(* IEC 61131-3 sources: ConveyorControl-with-PLC/4E_Gruppe1_Graf_Projekt1/Class/SafetyBase (part 5) *)

            // get state via SDO communication
            StandardRequest.SDOHeader.CRC  := 0;                                                   // CRC is always 0 in Std communication
            StandardRequest.SDOHeader.Cmd  := SB_SDO_COMMAND_GET_DIAG_INFO;                        // read command
            StandardRequest.SDOHeader.Typ  := SDO_STD;                                             // standard frame type
            StandardRequest.SDOHeader.SeqNr:= StandardSeqNr OR 16#80;                              // sequence number
            StandardRequest.SDOHeader.Len  := 4 + 1;                                               // header + µC-selection
            StandardRequest.aData[0] := DiagVars.ucChoiceDiagInfo;

            LastRequest := _DiagInfo;

#ifdef SAFETY_PROTOCOL_ANALYZER_ACTIVATED
  RecordFrame((#StandardRequest)$^DINT, 1);
#endif

            //copy SDO into write-buffer
            ToStdLib.MemCpy(dest := #p_Handle_SDO_Write^.SDOStructure, source := #StandardRequest, size := (sizeof(SDOHeader.StdHeader.CRC) + StandardRequest.SDOHeader.Len));

            //mark SDO data as valid
            p_Handle_SDO_Write^.us_Status := SAFETY_SDO_DATA_VALID;

            if ( pISafety^.udVersion >= 16#1001 ) then
              SAFETY_iPushSafetyTask();
            end_if;

          else

            if SchedulerStepNo = 6 then
              UnsafeScheduler := UnsafeSchedulerGetDiagVars;

            elsif SchedulerStepNo = 7 then
              UnsafeScheduler := UnsafeSchedulerGetRetryCounter;
            end_if;

          end_if;
       (* ***************************************** *)
          UnsafeSchedulerGetRetryCounter:
       (* ***************************************** *)
           //read out the retry counters every 10seconds
          if (ops.tAbsolute - ud_RetryCntTimeMark) > SB_RETRY_COUNTER_WAIT_TIME  then

            SDORequestBuffer.StdHeader.CRC  := 0;                                                         // CRC is always 0 in Std communication
            SDORequestBuffer.StdHeader.Cmd  := SB_SDO_COMMAND_READ;                                       // read command
            SDORequestBuffer.StdHeader.Typ  := SDO_STD;                                                   // standard frame type
            SDORequestBuffer.StdHeader.SeqNr:= StandardSeqNr OR 16#80;                                    // sequence number
            SDORequestBuffer.StdHeader.Len  := 4 + 4 + SB_SDO_LENGTH_RETRY_COUNTER;                       // header + destination address + length of data
            SDORequestBuffer.ud_Address     := SB_SDO_ADDRESS_RETRY_COUNTER;                              // address of retrycounter
            SDORequestBuffer.us_Length      := SB_SDO_LENGTH_RETRY_COUNTER;                               // length of data

            LastRequest := _ReadRetryCounter;

  #ifdef SAFETY_PROTOCOL_ANALYZER_ACTIVATED
  RecordFrame((#SDORequestBuffer)$^DINT, 1);
  #endif

            //copy SDO into write-buffer
            ToStdLib.MemCpy(dest := #p_Handle_SDO_Write^.SDOStructure, source := #SDORequestBuffer, size := (sizeof(SDOHeader.StdHeader.CRC) + SDORequestBuffer.StdHeader.Len));

            //mark SDO data as valid
            p_Handle_SDO_Write^.us_Status := SAFETY_SDO_DATA_VALID;

            if ( pISafety^.udVersion >= 16#1001 ) then
              SAFETY_iPushSafetyTask();
            end_if;

            //reset timemark
            ud_RetryCntTimeMark := ops.tAbsolute;

          else
            UnsafeScheduler := UnsafeSchedulerGetDiagVars;
          end_if;
        else
          LogError("Undefined Scheduler-State");
        end_case;
      end_while;
    end_if;
  end_if;

  // at the first run we write all variables independent of any changes
  if RunState > OldRunState then
    SendAllUnsafeValues();
  end_if;
  OldRunState := RunState;

	state := READY;

//============================ Profiler start======================================================
#ifdef  DM_Profiler
  StopTimeMeasurement(usMode := DMTIME_CY);
#endif
//============================ Profiler end========================================================
END_FUNCTION

FUNCTION SafetyBase::GetPointer2IFPDOBuffer
	VAR_OUTPUT
		ud_PDOBuffer 	: UDINT;
	END_VAR

  IFPDOOutputIsUsed := TRUE;

  //set pointer to address of buffer pointer
  ud_PDOBuffer := ( #IFPDOOutputBuffer )$UDINT;

END_FUNCTION

FUNCTION VIRTUAL SafetyBase::GetConfiguration

END_FUNCTION

FUNCTION SafetyBase::AddMovDOs
	VAR_OUTPUT
		ret_code 	: iprStates;
	END_VAR
  VAR
  	tempCmd         : CmdStruct;
    _result         : results;
    dataADDDO       : t_AddMoveDOCfg;
    i               : DINT;
  END_VAR

  ret_code := READY;

  // at the connect of the module we read the needed write size (written by the safety designer). at this point we know if the module needs data. if not => no move necessary
  if MyPDOWriteSize = 0 then
    return;
  end_if;

  // this stays the same for every DO
  tempCmd.uiCmd     := _BUS_IF_ADD_MOVE_DO;
  tempCmd.aPara[0]  := (#dataADDDO)$DINT;

  // initialize the parameter structure
  dataADDDO.ud_length_move        := MyPDOWriteSize;
  dataADDDO.ud_handle_source      := 0; // is set via SdiasManager or similar
  dataADDDO.ud_addressoff_source  := 0; // is set via SdiasManager or similar
  dataADDDO.p_sourcedata          := pPDOReadData;
  dataADDDO.ud_handle_dest        := 0; // is set via SdiasManager or similar
  dataADDDO.ud_addressoff_dest    := 0; // is set via SdiasManager or similar
  dataADDDO.p_destdata            := pPDOWriteData;
  dataADDDO.Priority              := _BUS_IF_ISO_MOVE;

  ToBusInterface.NewInst(pPara:=#tempCmd, pResult:=#_result);
  if _result.aData[0]$t_BusIFRetvalErrorcode = _BUS_IF_RETVAL_OK then
    InputMovSettings.MoveSettingsBusIF.Handle               := _result.aData$t_AddMoveDORet.Handle;
    InputMovSettings.MoveSettingsBusIF.ud_length_move       := dataADDDO.ud_length_move;
    InputMovSettings.MoveSettingsBusIF.ud_handle_source     := dataADDDO.ud_handle_source;
    InputMovSettings.MoveSettingsBusIF.ud_addressoff_source := dataADDDO.ud_addressoff_source;
    InputMovSettings.MoveSettingsBusIF.p_sourcedata         := dataADDDO.p_sourcedata;
    InputMovSettings.MoveSettingsBusIF.ud_handle_dest       := dataADDDO.ud_handle_dest;
    InputMovSettings.MoveSettingsBusIF.ud_addressoff_dest   := dataADDDO.ud_addressoff_dest;
    InputMovSettings.MoveSettingsBusIF.p_destdata           := dataADDDO.p_destdata;
    InputMovSettings.EnableState                            := _BUS_IF_RUN_STATE_NO_RUN;

    // addresses of local PDOs (set after creating the Move-DO, because we don't have the pointers to the DPRAM before (only in local memory)
    ud_LocalMoveSourceAddr := dataADDDO.p_sourcedata$UDINT;
    ud_LocalMoveDestAddr   := dataADDDO.p_destdata$UDINT;

    ud_LocalReadHandle     := dataADDDO.ud_handle_source;
    ud_LocalReadOffset     := dataADDDO.ud_addressoff_source;

    ud_LocalWriteHandle    := dataADDDO.ud_handle_dest;
    ud_LocalWriteOffset    := dataADDDO.ud_addressoff_dest;
  else
    LogError("(SafetyBase::AddMovDOs) Failed to add move DO");
    ret_code := ERROR;
  end_if;

  if (AdditionalSPDOs > 0) then
    for i := 0 to (AdditionalSPDOs-1) do
      dataADDDO.p_destdata  := aAdditionalPDOs[i].pPDOWriteData;

      ToBusInterface.NewInst(pPara:=#tempCmd, pResult:=#_result);
      if _result.aData[0]$t_BusIFRetvalErrorcode = _BUS_IF_RETVAL_OK then
        aAdditionalPDOs[i].InputMovSettings.MoveSettingsBusIF.Handle                := _result.aData$t_AddMoveDORet.Handle;
        aAdditionalPDOs[i].InputMovSettings.MoveSettingsBusIF.ud_length_move        := dataADDDO.ud_length_move;
        aAdditionalPDOs[i].InputMovSettings.MoveSettingsBusIF.ud_handle_source      := dataADDDO.ud_handle_source;
        aAdditionalPDOs[i].InputMovSettings.MoveSettingsBusIF.ud_addressoff_source  := dataADDDO.ud_addressoff_source;
        aAdditionalPDOs[i].InputMovSettings.MoveSettingsBusIF.p_sourcedata          := dataADDDO.p_sourcedata;
        aAdditionalPDOs[i].InputMovSettings.MoveSettingsBusIF.ud_handle_dest        := dataADDDO.ud_handle_dest;
        aAdditionalPDOs[i].InputMovSettings.MoveSettingsBusIF.ud_addressoff_dest    := dataADDDO.ud_addressoff_dest;
        aAdditionalPDOs[i].InputMovSettings.MoveSettingsBusIF.p_destdata            := dataADDDO.p_destdata;
        aAdditionalPDOs[i].InputMovSettings.EnableState                             := _BUS_IF_RUN_STATE_NO_RUN;

        aAdditionalPDOs[i].ud_LocalMoveDestAddr := dataADDDO.p_destdata$UDINT;
        aAdditionalPDOs[i].ud_LocalWriteHandle  := dataADDDO.ud_handle_dest$UDINT;
        aAdditionalPDOs[i].ud_LocalWriteOffset  := dataADDDO.ud_addressoff_dest$UDINT;
      else
        LogError("(SafetyBase::AddMovDOs) Failed to add move DO for additional write PDOs");
        ret_code := ERROR;
      end_if;
    end_for;
  end_if;

  // now get the access info needed for the move command
  tempCmd.uiCmd     := _BUS_IF_GET_ACCESS_INFO;
  tempCmd.aPara[0]  := pPDOIFReadData$DINT;

  ToBusInterface.NewInst(pPara:=#tempCmd, pResult:=#_result);
  if _result.aData[0]$t_AccessInfoRet.retcode = _BUS_IF_RETVAL_OK then
    ud_LocalMoveIFSourceAddr  := (_result.aData[0]$t_AccessInfoRet.p_dataDPRAM)$HDINT;
    ud_LocalIFReadHandle      := _result.aData[0]$t_AccessInfoRet.ud_handle;
    ud_LocalIFReadOffset      := _result.aData[0]$t_AccessInfoRet.ud_addressoff;
  else
    LogError("(SafetyBase::AddMovDOs) Failed to get access info for interface read access");
    ret_code := ERROR;
  end_if;

  b_MoveDOsCreated := TRUE;

END_FUNCTION

FUNCTION SafetyBase::UpdateMovDO
	VAR_INPUT
		p_MoveSettings 	: ^t_MoveSettings;
		ud_NewSourceHandle 	: UDINT;
		ud_NewSourceOffset 	: UDINT;
		ud_NewSourcePointer 	: UDINT;
		ui_NewLength 	: UINT;
	END_VAR
  VAR
  	b_DifferenceDetected : BOOL;
  	tempCmd         : CmdStruct;
    _result         : results;
  END_VAR

  // check if there is a difference to the old settings
  b_DifferenceDetected := FALSE;

  if ud_NewSourceHandle <> p_MoveSettings^.MoveSettingsBusIF.ud_handle_source then
    p_MoveSettings^.MoveSettingsBusIF.ud_handle_source := ud_NewSourceHandle;
    b_DifferenceDetected := TRUE;
  end_if;

  if ud_NewSourceOffset <> p_MoveSettings^.MoveSettingsBusIF.ud_addressoff_source then
    p_MoveSettings^.MoveSettingsBusIF.ud_addressoff_source := ud_NewSourceOffset;
    b_DifferenceDetected := TRUE;
  end_if;

  if ud_NewSourcePointer <> p_MoveSettings^.MoveSettingsBusIF.p_sourcedata$UDINT then
    p_MoveSettings^.MoveSettingsBusIF.p_sourcedata$UDINT := ud_NewSourcePointer;
    b_DifferenceDetected := TRUE;
  end_if;

  if ui_NewLength <> p_MoveSettings^.MoveSettingsBusIF.ud_length_move then
    p_MoveSettings^.MoveSettingsBusIF.ud_length_move := ui_NewLength;
    b_DifferenceDetected := TRUE;
  end_if;

  // if there is a difference to the old settings => change the move DO
  if b_DifferenceDetected then
    tempCmd.uiCmd     := _BUS_IF_UPDATE_MOVE_DO;
    tempCmd.aPara[0]  := (#p_MoveSettings^.MoveSettingsBusIF)$DINT;

    ToBusInterface.NewInst(pPara:=#tempCmd, pResult:=#_result);
    if _result.aData[0]$t_BusIFRetvalErrorcode <> _BUS_IF_RETVAL_OK then
      LogError("(SafetyBase::UpdateMovDO) Failed to change move-DO");
    end_if;
  end_if;

  // if the Move-DO is'nt started
  if p_MoveSettings^.EnableState <> _BUS_IF_RUN_STATE_CONT_RUN then
    // => start it, because we have to move in every cycle
    SetDORunState(Handle := p_MoveSettings^.MoveSettingsBusIF.Handle, NewState:=_BUS_IF_RUN_STATE_CONT_RUN);
    p_MoveSettings^.EnableState := _BUS_IF_RUN_STATE_CONT_RUN;
  end_if;

END_FUNCTION

FUNCTION VIRTUAL SafetyBase::SetSafetyState
	VAR_INPUT
		NewState 	: SafetyConfigStateType;
	END_VAR

  // use it locally => can also be forwarded in derivation
  SafetyState := NewState;

END_FUNCTION

FUNCTION VIRTUAL SafetyBase::RefreshAsySrv
  // derive this
END_FUNCTION

FUNCTION VIRTUAL SafetyBase::SetRetryCounter

  SafetyRetryCounter := -1;

END_FUNCTION

FUNCTION SafetyBase::IsInCache
	VAR_INPUT
		ud_Address 	: UDINT;
		us_Length 	: USINT;
	END_VAR
	VAR_OUTPUT
		ItsInside 	: BOOL;
	END_VAR

  if CachedSize &
     (ud_Address >= CachedAddr) &
     ((ud_Address + us_Length) <= (CachedAddr + CachedSize)) then
    ItsInside := TRUE;
  else
    ItsInside := FALSE;
  end_if;

END_FUNCTION

FUNCTION SafetyBase::AddToCache
	VAR_INPUT
		p_SDORequestBuffer 	: ^SDORequReadConfig;
		p_SDOResponseBuffer 	: ^SDORespReadConfig;
	END_VAR

  if p_SDORequestBuffer^.us_Length then
    CachedAddr := p_SDORequestBuffer^.ud_Address;
    CachedSize := p_SDORequestBuffer^.us_Length;
    _memcpy(ptr1:=#Cache, ptr2:=#p_SDOResponseBuffer^.ud_Data, cntr:=p_SDORequestBuffer^.us_Length);
  end_if;

END_FUNCTION
